(*
SPDX-FileCopyrightText: © 2026 Oleksandr Tiutyk <trofimich@gmail.com>
SPDX-License-Identifier: MIT
License: https://opensource.org/license/mit
*)

(*!
<summary>Provides fluent assertions on a copied BOOL value.</summary>
<description>
Copies actual into persistent instance storage before the entry method returns; literals and expression
results therefore remain valid throughout the immediate chain. Owns no heap allocation or pointed-to resource.
The message prefixes every failure until the next preparation. Finish one chain before starting another on
the owning Assertions provider. Use only from the owning test callback on one task, without reentry.
Obtain this context from the owning provider; direct unprepared use is unsupported.
Expected arguments use the declared IEC type; ordinary compiler conversions happen before comparison.
This context does not depend on another assertion context.
Object metadata is available before preparation; inherited equality compares instance identity.
</description>
*)

{attribute 'no_explicit_call' := 'do not call this function block directly'}
FUNCTION_BLOCK BoolAssertionContext EXTENDS TOF_Core.Object
VAR_STAT
	{attribute 'hide'}
	_ClassName : STRING := __POUNAME();
END_VAR
VAR
	_Actual : BOOL;
	_TestCase : ITestCase;
	_Message : WSTRING(255);
END_VAR

(*!
<summary>Provides the implementation class name.</summary>
<description>
Borrowed read-only reference to compiler-initialized storage, valid throughout the instance lifetime.
Do not modify the returned reference; no ownership is transferred.
</description>
*)
{attribute 'monitoring' := 'call'}
PROPERTY ClassName : REFERENCE TO STRING
GET
ClassName REF= _ClassName;
END_GET
END_PROPERTY

(*!
<summary>Asserts that the actual Boolean value is FALSE.</summary>
<description>
Records failure without interrupting the callback; preserves the chain message.
</description>
*)
METHOD FINAL IsFalse : REFERENCE TO BoolAssertionContext
IF _Actual THEN
	failComparison(expected := FALSE, expectation := "Expected: ");
END_IF

IsFalse REF= THIS^;
END_METHOD

(*!
<summary>Asserts that the actual Boolean value is TRUE.</summary>
<description>
Records failure without interrupting the callback; preserves the chain message.
</description>
*)
METHOD FINAL IsTrue : REFERENCE TO BoolAssertionContext
IF NOT _Actual THEN
	failComparison(expected := TRUE, expectation := "Expected: ");
END_IF

IsTrue REF= THIS^;
END_METHOD

(*!
<summary>Provides the library namespace.</summary>
<description>
Borrowed read-only reference to the compiler-initialized namespace, valid throughout the instance lifetime.
Do not modify the returned reference; no ownership is transferred.
</description>
*)
{attribute 'monitoring' := 'call'}
PROPERTY NamespaceName : REFERENCE TO STRING
GET
NamespaceName REF= CurrentNamespace.Name;
END_GET
END_PROPERTY

(*!
<summary>Asserts inequality with the expected value.</summary>
<description>
Records failure without interrupting the callback; preserves the message for the rest of the chain.
</description>
<param name="expected">Expected value converted by the compiler to BOOL.</param>
*)
METHOD FINAL NotToBe : REFERENCE TO BoolAssertionContext
VAR_INPUT
	expected : BOOL;
END_VAR
IF _Actual = expected THEN
	failComparison(
		expected := expected,
		expectation := "Expected value not to be: "
	);
END_IF

NotToBe REF= THIS^;
END_METHOD

(*!
<summary>Copies the actual operand and replaces the chain-wide message.</summary>
<description>
Called by the owning Assertions provider after it verifies the running test case.
No pointer to this method's input storage is retained. The receiver is borrowed until the next preparation;
the owning provider keeps it alive throughout the immediate chain.
</description>
<param name="actual">Value copied into this context.</param>
<param name="testCase">Borrowed failure receiver for the immediate chain.</param>
<param name="message">Copied diagnostic prefix, including empty to clear the previous prefix.</param>
*)
METHOD INTERNAL FINAL Prepare
VAR_INPUT
	actual : BOOL;
	testCase : ITestCase;
END_VAR
VAR_IN_OUT CONSTANT
	message : WSTRING(255);
END_VAR
_Actual := actual;
_TestCase := testCase;
_Message := message;
END_METHOD

(*!
<summary>Reports the byte size of this concrete instance.</summary>
<description>
Includes inline fields and nested instances, but excludes separately allocated payloads.
Obtaining the size does not transfer ownership or validate an arbitrary address.
</description>
*)
{attribute 'monitoring' := 'call'}
PROPERTY SelfSize : ULINT
GET
SelfSize := XSIZEOF(THIS^);
END_GET
END_PROPERTY

(*!
<summary>Asserts equality with the expected value.</summary>
<description>
Records failure without interrupting the callback; preserves the message for the rest of the chain.
</description>
<param name="expected">Expected value converted by the compiler to BOOL.</param>
*)
METHOD FINAL ToBe : REFERENCE TO BoolAssertionContext
VAR_INPUT
	expected : BOOL;
END_VAR
IF _Actual <> expected THEN
	failComparison(
		expected := expected,
		expectation := "Expected: "
	);
END_IF

ToBe REF= THIS^;
END_METHOD

(*!
<summary>Formats a failed typed predicate and reports it with the chain message.</summary>
<description>
Does not change operands or chain state. The receiver retains its first failure. Reporting exceptions
propagate to the enclosing test callback handler; an unprepared receiver is a configuration error.
</description>
<param name="expected">Typed expected operand used only for this diagnostic.</param>
<param name="expectation">Prefix identifying the failed predicate.</param>
*)
METHOD PRIVATE failComparison
VAR_INPUT
	expected : BOOL;
	expectation : WSTRING(40);
END_VAR
VAR
	actualText : WSTRING(255);
	expectedText : WSTRING(255);
	diagnostic : TOF_Core.ERROR_MESSAGE;
END_VAR
actualText := TO_WSTRING(_Actual);
expectedText := TO_WSTRING(expected);

diagnostic := TOF_Core.WideStrings.Concat255(
	expectation,
	expectedText,
	", but was: ",
	actualText
);

TestServices.ReportAssertionFailure(
	testCase := _TestCase,
	message := _Message,
	sourceClassName := ClassName,
	defaultMessage := diagnostic
);
END_METHOD

END_FUNCTION_BLOCK

(* stored: Version 1.1.0.1
   POU BoolAssertionContext: Id {efe27691-50c3-4b7d-8d0b-f55e2e145187}, SpecialFunc None
   Folder Service methods: Id {7b71b26c-d44d-49f6-a850-725fe7b9ef2d}
   Property ClassName: Id {4ca1faa7-e905-4b69-9307-351b17a85f6e}
   Get Get: Id {3324de6b-4837-4938-a01a-7157edbd7e3e}
   Method IsFalse: Id {1543e475-9b31-499a-80e9-413ce53c0daf}
   Method IsTrue: Id {fbe114fd-1da5-4b3f-834b-963b6c1e02ce}
   Property NamespaceName: Id {62cf25de-65d4-47ae-a57c-558483847e71}
   Get Get: Id {79e4332a-d5c7-4dda-83fa-27d6cd93ce8e}
   Method NotToBe: Id {eb9f27c6-e501-4e76-b75a-a8a3c88d029f}
   Method Prepare: Id {4a74021a-f6cb-410a-8374-f2fbbcb24a04}
   Property SelfSize: Id {8961f7b7-72bd-4b81-84dd-c2a2e2fd695d}
   Get Get: Id {5024db69-413b-4043-b6ff-da3c843390cd}
   Method ToBe: Id {947bbb76-d07b-440b-8b47-e242c2dbc887}
   Method failComparison: Id {f823a0f6-77e1-4d52-8453-5ab1096f607a} *)
